Fanuc KAREL source: KB00201.KL

PROGRAM KB00201
%NOLOCKGROUP
VAR
  P1: FILE
  P2: STRING[80]
  P3: INTEGER
  P4: INTEGER
BEGIN
  P2 = 'A'
  P3 = 1
  P4 = 1
  XML_SCAN(P1, P2, P3, P4)
END KB00201
